// TIA Portal V19 export
DATA_BLOCK "MCP_RC_DB2"   // DB9802
{ S7_Optimized_Access := 'TRUE' }
   VAR
      Count : Int := 5;
      Motor : "MCP_RC_UDT";
   END_VAR
BEGIN
END_DATA_BLOCK
